// TIA Portal V20 export
DATA_BLOCK "05_Not-Aus_DB"   // DB164
// stored: InstanceOfName 05_Not-Aus, InstanceOfType FB
"05_Not-Aus"
BEGIN
END_DATA_BLOCK
